(* IEC 61131-3 sources: plcassist-cli/packages/volt-lsp-iec/test-corpus/pro2193/Device/Plc Logic/Application/09 Misc/Library Manager/SysSocket Implementation, 44 files *)

(* ---- SYSSOCKACCEPT.fun ---- *)
FUNCTION SYSSOCKACCEPT : RTS_IEC_HANDLE
VAR_INPUT
	HSOCKET : RTS_IEC_HANDLE;
	PSOCKADDR : POINTER TO SOCKADDRESS;
	PDISOCKADDRSIZE : POINTER TO DINT;
	PRESULT : POINTER TO RTS_IEC_RESULT;
END_VAR
END_FUNCTION

(* ---- SYSSOCKBIND.fun ---- *)
FUNCTION SYSSOCKBIND : RTS_IEC_RESULT
VAR_INPUT
	HSOCKET : RTS_IEC_HANDLE;
	PSOCKADDR : POINTER TO SOCKADDRESS;
	DISOCKADDRSIZE : DINT;
END_VAR
END_FUNCTION

(* ---- SYSSOCKCLOSE.fun ---- *)
FUNCTION SYSSOCKCLOSE : RTS_IEC_RESULT
VAR_INPUT
	HSOCKET : RTS_IEC_HANDLE;
END_VAR
END_FUNCTION

(* ---- SYSSOCKCLOSEUDP.fun ---- *)
FUNCTION SYSSOCKCLOSEUDP : RTS_IEC_RESULT
VAR_INPUT
	HSOCKETUDP : RTS_IEC_HANDLE;
END_VAR
END_FUNCTION

(* ---- SYSSOCKCONNECT.fun ---- *)
FUNCTION SYSSOCKCONNECT : RTS_IEC_RESULT
VAR_INPUT
	HSOCKET : RTS_IEC_HANDLE;
	PSOCKADDR : POINTER TO SOCKADDRESS;
	DISOCKADDRSIZE : DINT;
END_VAR
END_FUNCTION

(* ---- SYSSOCKCREATE.fun ---- *)
FUNCTION SYSSOCKCREATE : RTS_IEC_HANDLE
VAR_INPUT
	IADDRESSFAMILY : INT;
	DITYPE : DINT;
	DIPROTOCOL : DINT;
	PRESULT : POINTER TO RTS_IEC_RESULT;
END_VAR
END_FUNCTION

(* ---- SYSSOCKCREATEUDP.fun ---- *)
FUNCTION SYSSOCKCREATEUDP : RTS_IEC_HANDLE
VAR_INPUT
	DISENDPORT : DINT;
	DIRECVPORT : DINT;
	PRESULT : POINTER TO RTS_IEC_RESULT;
END_VAR
END_FUNCTION

(* ---- SYSSOCKFDINIT.fun ---- *)
FUNCTION SYSSOCKFDINIT : RTS_IEC_RESULT
VAR_INPUT
	HSOCKET : RTS_IEC_HANDLE;
	PFS : REFERENCE TO SOCKET_FD_SET;
END_VAR
END_FUNCTION

(* ---- SYSSOCKFDISSET.fun ---- *)
FUNCTION SYSSOCKFDISSET : BOOL
VAR_INPUT
	HSOCKET : RTS_IEC_HANDLE;
	PFS : REFERENCE TO SOCKET_FD_SET;
END_VAR
END_FUNCTION

(* ---- SYSSOCKFDZERO.fun ---- *)
FUNCTION SYSSOCKFDZERO : RTS_IEC_RESULT
VAR_INPUT
	PFS : REFERENCE TO SOCKET_FD_SET;
END_VAR
END_FUNCTION

(* ---- SYSSOCKGETFIRSTADAPTERINFO.fun ---- *)
FUNCTION SYSSOCKGETFIRSTADAPTERINFO : RTS_IEC_HANDLE
VAR_INPUT
	PADAPTERINFO : POINTER TO SOCK_ADAPTER_INFORMATION;
	PUXIADAPTERINFOSIZE : POINTER TO __UXINT;
	PRESULT : POINTER TO RTS_IEC_RESULT;
END_VAR
END_FUNCTION

(* ---- SYSSOCKGETHOSTBYNAME.fun ---- *)
FUNCTION SYSSOCKGETHOSTBYNAME : RTS_IEC_RESULT
VAR_INPUT
	SZHOSTNAME : REFERENCE TO STRING;
	PHOST : POINTER TO SOCK_HOSTENT;
END_VAR
END_FUNCTION

(* ---- SYSSOCKGETHOSTNAME.fun ---- *)
FUNCTION SYSSOCKGETHOSTNAME : RTS_IEC_RESULT
VAR_INPUT
	SZHOSTNAME : REFERENCE TO STRING;
	DINAMELEN : DINT;
END_VAR
END_FUNCTION

(* ---- SYSSOCKGETNEXTADAPTERINFO.fun ---- *)
FUNCTION SYSSOCKGETNEXTADAPTERINFO : RTS_IEC_HANDLE
VAR_INPUT
	HPREVADAPTER : RTS_IEC_HANDLE;
	PADAPTERINFO : POINTER TO SOCK_ADAPTER_INFORMATION;
	PUXIADAPTERINFOSIZE : POINTER TO __UXINT;
	PRESULT : POINTER TO RTS_IEC_RESULT;
END_VAR
END_FUNCTION

(* ---- SYSSOCKGETOPTION.fun ---- *)
FUNCTION SYSSOCKGETOPTION : RTS_IEC_RESULT
VAR_INPUT
	HSOCKET : RTS_IEC_HANDLE;
	DILEVEL : DINT;
	DIOPTION : DINT;
	PDIOPTIONVALUE : POINTER TO DINT;
	PDIOPTIONLEN : POINTER TO DINT;
END_VAR
END_FUNCTION

(* ---- SYSSOCKGETOSHANDLE.fun ---- *)
FUNCTION SYSSOCKGETOSHANDLE : RTS_IEC_HANDLE
VAR_INPUT
	HSOCKETUDP : RTS_IEC_HANDLE;
END_VAR
END_FUNCTION

(* ---- SYSSOCKGETPEERNAME.fun ---- *)
FUNCTION SYSSOCKGETPEERNAME : RTS_IEC_RESULT
VAR_INPUT
	HSOCKET : RTS_IEC_HANDLE;
	PSOCKADDR : POINTER TO SOCKADDRESS;
	PDISOCKADDRSIZE : POINTER TO DINT;
END_VAR
END_FUNCTION

(* ---- SYSSOCKGETRECVSIZEUDP.fun ---- *)
FUNCTION SYSSOCKGETRECVSIZEUDP : __XINT
VAR_INPUT
	HSOCKETUDP : RTS_IEC_HANDLE;
	DITIMEOUT : DINT;
	PRESULT : POINTER TO RTS_IEC_RESULT;
END_VAR
END_FUNCTION

(* ---- SYSSOCKGETSOCKNAME.fun ---- *)
FUNCTION SYSSOCKGETSOCKNAME : RTS_IEC_RESULT
VAR_INPUT
	HSOCKET : RTS_IEC_HANDLE;
	PSOCKADDR : POINTER TO SOCKADDRESS;
	PDISOCKADDRSIZE : POINTER TO DINT;
END_VAR
END_FUNCTION

(* ---- SYSSOCKGETSUBNETMASK.fun ---- *)
FUNCTION SYSSOCKGETSUBNETMASK : RTS_IEC_RESULT
VAR_INPUT
	SZIPADDRESS : REFERENCE TO STRING;
	SZSUBNETMASK : REFERENCE TO STRING;
	DIMAXSUGNETMASK : DINT;
END_VAR
END_FUNCTION

(* ---- SYSSOCKHTONL.fun ---- *)
FUNCTION SYSSOCKHTONL : UDINT
VAR_INPUT
	ULHOST : UDINT;
END_VAR
END_FUNCTION

(* ---- SYSSOCKHTONS.fun ---- *)
FUNCTION SYSSOCKHTONS : WORD
VAR_INPUT
	USHOST : WORD;
END_VAR
END_FUNCTION

(* ---- SYSSOCKINETADDR.fun ---- *)
FUNCTION SYSSOCKINETADDR : RTS_IEC_RESULT
VAR_INPUT
	SZIPADDRESS : REFERENCE TO STRING;
	PINADDR : POINTER TO UDINT;
END_VAR
END_FUNCTION

(* ---- SYSSOCKINETNTOA.fun ---- *)
FUNCTION SYSSOCKINETNTOA : RTS_IEC_RESULT
VAR_INPUT
	PINADDR : POINTER TO INADDR;
	SZIPADDR : REFERENCE TO STRING;
	DIIPADDRSIZE : DINT;
END_VAR
END_FUNCTION

(* ---- SYSSOCKIOCTL.fun ---- *)
FUNCTION SYSSOCKIOCTL : RTS_IEC_RESULT
VAR_INPUT
	HSOCKET : RTS_IEC_HANDLE;
	DICOMMAND : DINT;
	PDIPARAMETER : POINTER TO DINT;
END_VAR
END_FUNCTION

(* ---- SYSSOCKLISTEN.fun ---- *)
FUNCTION SYSSOCKLISTEN : RTS_IEC_RESULT
VAR_INPUT
	HSOCKET : RTS_IEC_HANDLE;
	DIMAXCONNECTIONS : DINT;
END_VAR
END_FUNCTION

(* ---- SYSSOCKNTOHL.fun ---- *)
FUNCTION SYSSOCKNTOHL : UDINT
VAR_INPUT
	ULNET : UDINT;
END_VAR
END_FUNCTION

(* ---- SYSSOCKNTOHS.fun ---- *)
FUNCTION SYSSOCKNTOHS : WORD
VAR_INPUT
	USNET : WORD;
END_VAR
END_FUNCTION

(* ---- SYSSOCKPING.fun ---- *)
FUNCTION SYSSOCKPING : RTS_IEC_RESULT
VAR_INPUT
	SZIPADDRESS : REFERENCE TO STRING;
	ULTIMEOUT : UDINT;
	PULREPLYTIME : POINTER TO UDINT;
END_VAR
END_FUNCTION

(* ---- SYSSOCKRECV.fun ---- *)
FUNCTION SYSSOCKRECV : __XINT
VAR_INPUT
	HSOCKET : RTS_IEC_HANDLE;
	PBYBUFFER : POINTER TO BYTE;
	DIBUFFERSIZE : __XINT;
	DIFLAGS : DINT;
	PRESULT : POINTER TO RTS_IEC_RESULT;
END_VAR
END_FUNCTION

(* ---- SYSSOCKRECVFROM.fun ---- *)
FUNCTION SYSSOCKRECVFROM : __XINT
VAR_INPUT
	HSOCKET : RTS_IEC_HANDLE;
	PBYBUFFER : POINTER TO BYTE;
	DIBUFFERSIZE : __XINT;
	DIFLAGS : DINT;
	PSOCKADDR : POINTER TO SOCKADDRESS;
	DISOCKADDRSIZE : DINT;
	PRESULT : POINTER TO RTS_IEC_RESULT;
END_VAR
END_FUNCTION

(* ---- SYSSOCKRECVFROMUDP.fun ---- *)
FUNCTION SYSSOCKRECVFROMUDP : __XINT
VAR_INPUT
	HSOCKETUDP : RTS_IEC_HANDLE;
	PBYDATA : POINTER TO BYTE;
	DIDATASIZE : __XINT;
	PREPLY : POINTER TO UDP_REPLY;
	PRESULT : POINTER TO RTS_IEC_RESULT;
END_VAR
END_FUNCTION

(* ---- SYSSOCKRECVFROMUDP2.fun ---- *)
FUNCTION SYSSOCKRECVFROMUDP2 : __XINT
VAR_INPUT
	HSOCKETUDP : RTS_IEC_HANDLE;
	PBYDATA : POINTER TO BYTE;
	DIDATASIZE : __XINT;
	PREPLY : POINTER TO UDP_REPLY2;
	PRESULT : POINTER TO RTS_IEC_RESULT;
END_VAR
END_FUNCTION

(* ---- SYSSOCKRECVMSG.fun ---- *)
FUNCTION SYSSOCKRECVMSG : __XINT
VAR_INPUT
	HSOCKET : RTS_IEC_HANDLE;
	PMESSAGE : POINTER TO SOCK_RECVMSG_MSG;
	FLAGS : DWORD;
	PRESULT : POINTER TO RTS_IEC_RESULT;
END_VAR
END_FUNCTION

(* ---- SYSSOCKSELECT.fun ---- *)
FUNCTION SYSSOCKSELECT : RTS_IEC_RESULT
VAR_INPUT
	DIWIDTH : DINT;
	PFDREAD : POINTER TO SOCKET_FD_SET;
	PFDWRITE : POINTER TO SOCKET_FD_SET;
	PFDEXCEPT : POINTER TO SOCKET_FD_SET;
	PTVTIMEOUT : POINTER TO SOCKET_TIMEVAL;
	PDIREADY : POINTER TO DINT;
END_VAR
END_FUNCTION

(* ---- SYSSOCKSEND.fun ---- *)
FUNCTION SYSSOCKSEND : __XINT
VAR_INPUT
	HSOCKET : RTS_IEC_HANDLE;
	PBYBUFFER : POINTER TO BYTE;
	DIBUFFERSIZE : __XINT;
	DIFLAGS : DINT;
	PRESULT : POINTER TO RTS_IEC_RESULT;
END_VAR
END_FUNCTION

(* ---- SYSSOCKSENDTO.fun ---- *)
FUNCTION SYSSOCKSENDTO : __XINT
VAR_INPUT
	HSOCKET : RTS_IEC_HANDLE;
	PBYBUFFER : POINTER TO BYTE;
	DIBUFFERSIZE : __XINT;
	DIFLAGS : DINT;
	PSOCKADDR : POINTER TO SOCKADDRESS;
	DISOCKADDRSIZE : DINT;
	PRESULT : POINTER TO RTS_IEC_RESULT;
END_VAR
END_FUNCTION

(* ---- SYSSOCKSENDTOUDP.fun ---- *)
FUNCTION SYSSOCKSENDTOUDP : __XINT
VAR_INPUT
	HSOCKETUDP : RTS_IEC_HANDLE;
	DIPORT : DINT;
	SZDESTADDRESS : REFERENCE TO STRING;
	PBYDATA : POINTER TO BYTE;
	DIDATASIZE : __XINT;
	PRESULT : POINTER TO RTS_IEC_RESULT;
END_VAR
END_FUNCTION

(* ---- SYSSOCKSETDEFAULTGATEWAY.fun ---- *)
FUNCTION SYSSOCKSETDEFAULTGATEWAY : RTS_IEC_RESULT
VAR_INPUT
	WSADAPTERNAME : REFERENCE TO WSTRING;
	GATEWAYADDR : REFERENCE TO INADDR;
END_VAR
END_FUNCTION

(* ---- SYSSOCKSETIPADDRESS.fun ---- *)
FUNCTION SYSSOCKSETIPADDRESS : RTS_IEC_RESULT
VAR_INPUT
	SZCARD : REFERENCE TO STRING;
	SZIPADDRESS : REFERENCE TO STRING;
END_VAR
END_FUNCTION

(* ---- SYSSOCKSETIPADDRESSANDNETMASK.fun ---- *)
FUNCTION SYSSOCKSETIPADDRESSANDNETMASK : RTS_IEC_RESULT
VAR_INPUT
	WSADAPTERNAME : REFERENCE TO WSTRING;
	IPADDR : REFERENCE TO INADDR;
	NETMASK : REFERENCE TO INADDR;
END_VAR
END_FUNCTION

(* ---- SYSSOCKSETOPTION.fun ---- *)
FUNCTION SYSSOCKSETOPTION : RTS_IEC_RESULT
VAR_INPUT
	HSOCKET : RTS_IEC_HANDLE;
	DILEVEL : DINT;
	DIOPTION : DINT;
	PDIOPTIONVALUE : POINTER TO DINT;
	DIOPTIONLEN : DINT;
END_VAR
END_FUNCTION

(* ---- SYSSOCKSETSUBNETMASK.fun ---- *)
FUNCTION SYSSOCKSETSUBNETMASK : RTS_IEC_RESULT
VAR_INPUT
	SZIPADDRESS : REFERENCE TO STRING;
	SZSUBNETMASK : REFERENCE TO STRING;
END_VAR
END_FUNCTION

(* ---- SYSSOCKSHUTDOWN.fun ---- *)
FUNCTION SYSSOCKSHUTDOWN : RTS_IEC_RESULT
VAR_INPUT
	HSOCKET : RTS_IEC_HANDLE;
	DIHOW : DINT;
END_VAR
END_FUNCTION
